TYPE ST_HW_DI :
STRUCT
END_STRUCT
END_TYPE

(* stored: Version 1.1.0.1, ProductVersion 3.1.4024.13
   DUT ST_HW_DI: Id {0cc95820-634c-4cca-bf0b-cea5000e8d43} *)
